Fanuc KAREL source: kf00117.KL

-- PROVISIONAL review KL for V940-1; original PC SHA256 7ccc8cfe116c08cdf244d07016f1a5b7941fa5f97f6ef0dc042e04593f1a6521
-- Incomplete behavior may be omitted. Consult companion uncertainty JSON. Do not deploy.
PROGRAM KF00117
%NOLOCKGROUP
BEGIN
  -- V9_ZERO_TABLE_METADATA_HINT layout=0001; no indexed target words; source/name/runtime held
  -- UNRESOLVED_PC offsets 0-1; opcodes 7B
  -- UNRESOLVED_PC offsets 6-21; opcodes 17,9D,33,34,23
  -- UNRESOLVED_PC offsets 26-30; opcodes 7F
  -- UNRESOLVED_PC offsets 35-45; opcodes 27,22,AA
  -- UNRESOLVED_PC offsets 50-54; opcodes 7F
END KF00117
